Staubli VAL3: zoneTemplate.dtx

public pointRx pO = {fatherId=world[0]}
public pointRx pX = {fatherId=world[0]}
public pointRx pY = {fatherId=world[0]}
public frame fBase = {fatherId=world[0]}
public pointRx pFirst = {fatherId=fBase[0]}
public pointRx pSecond = {fatherId=fBase[0]}
public bool bActive
public string sID
